VISUALIZATION Visu1  // 2x2
END_VISUALIZATION

(* stored: Version 1.1.0.1, ProductVersion 3.1.4026.0
   Visu Visu1: Id {a1b2c3d4-0000-0000-0000-000000000001} *)
